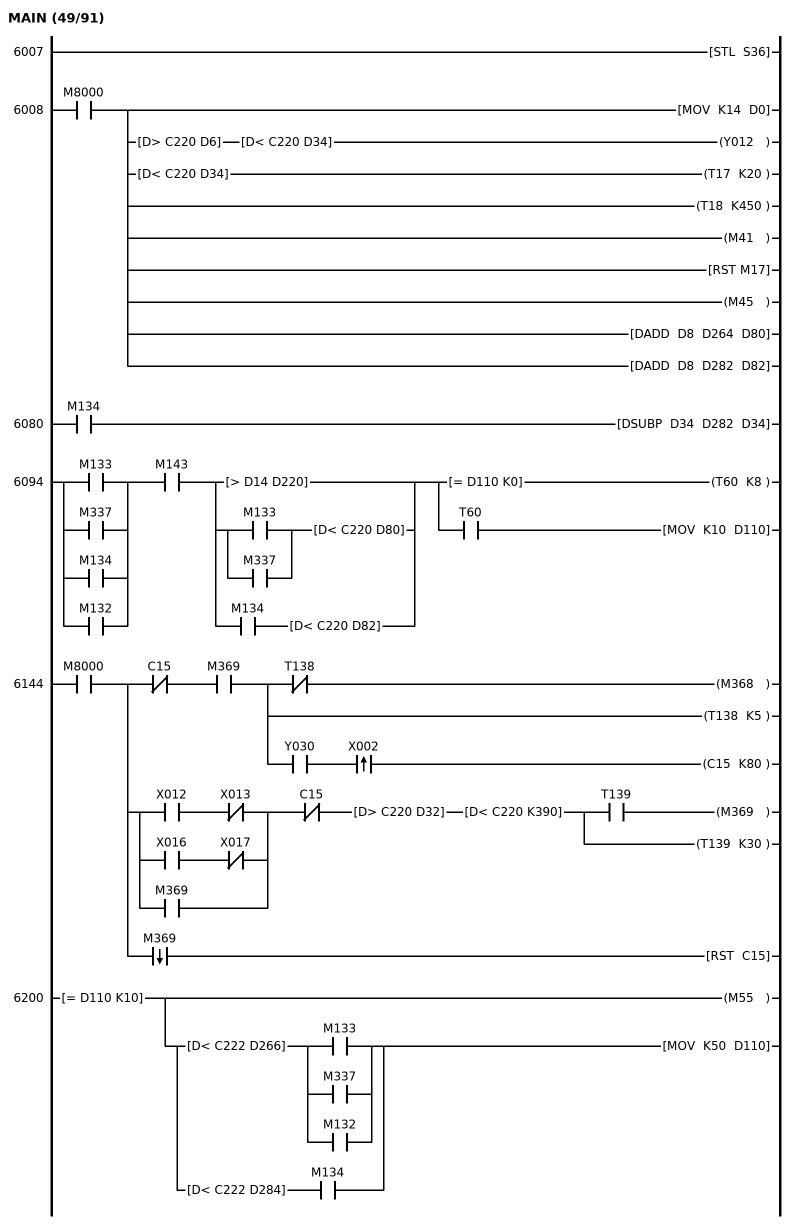
[picture p48: ladder of MAIN, rungs at steps 6007 to 6200]
6007  STL     S36
6008  LD      M8000
      MOV     K14 D0
      MPS
      ANDD>   C220 D6
      ANDD<   C220 D34
      OUT     Y012
      MRD
      ANDD<   C220 D34
      OUT     T17 K20
      MPP
      OUT     T18 K450
      OUT     M41
      RST     M17
      OUT     M45
      DADD    D8 D264 D80
      DADD    D8 D282 D82
6080  LD      M134
      DSUBP   D34 D282 D34
6094  LD      M133
      OR      M337
      OR      M134
      OR      M132
      AND     M143
      LD>     D14 D220
      LD      M133
      OR      M337
      ANDD<   C220 D80
      ORB
      LD      M134
      ANDD<   C220 D82
      ORB
      ANB
      MPS
      AND=    D110 K0
      OUT     T60 K8
      MPP
      AND     T60
      MOV     K10 D110
6144  LD      M8000
      MPS
      ANI     C15
      AND     M369
      MPS
      ANI     T138
      OUT     M368
      MPP
      OUT     T138 K5
      AND     Y030
      ANDP    X002
      OUT     C15 K80
      MRD
      LD      X012
      ANI     X013
      LD      X016
      ANI     X017
      ORB
      OR      M369
      ANB
      ANI     C15
      ANDD>   C220 D32
      ANDD<   C220 K390
      MPS
      AND     T139
      OUT     M369
      MPP
      OUT     T139 K30
      MPP
      ANDF    M369
      RST     C15
6200  LD=     D110 K10
      OUT     M55
      LDD<    C222 D266
      LD      M133
      OR      M337
      OR      M132
      ANB
      LDD<    C222 D284
      AND     M134
      ORB
      ANB
      MOV     K50 D110
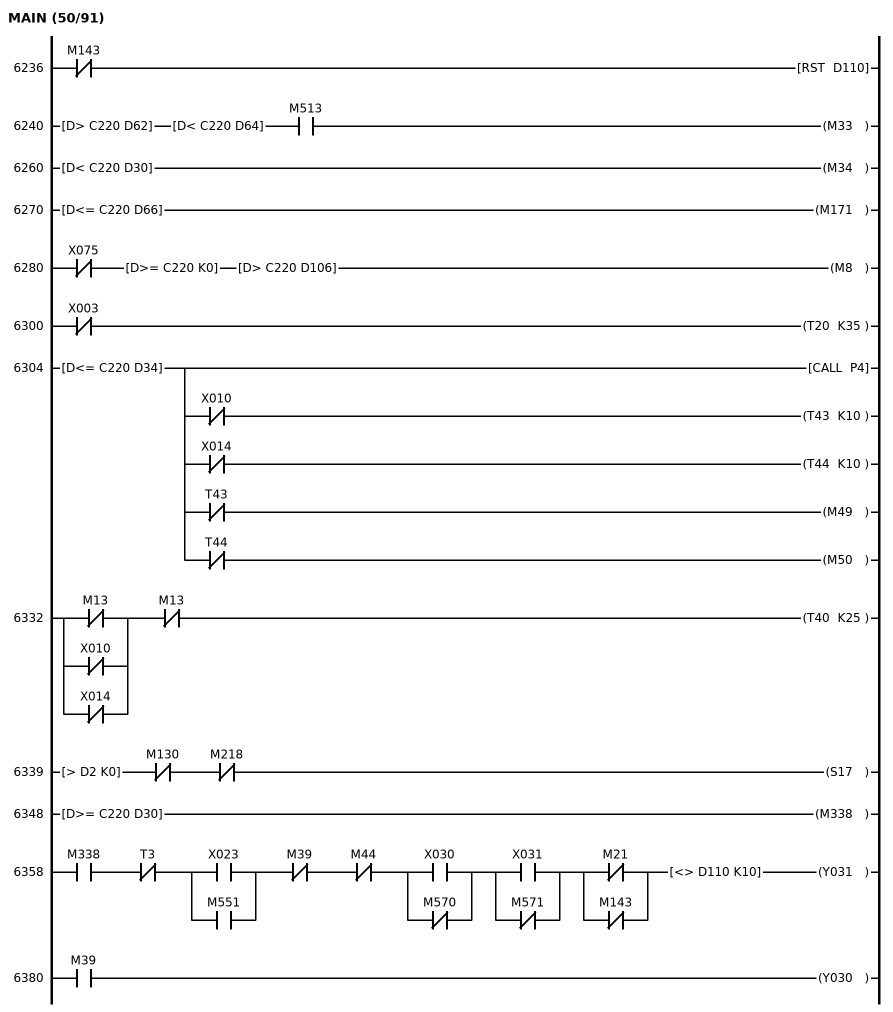
6236  LDI     M143
      RST     D110
6240  LDD>    C220 D62
      ANDD<   C220 D64
      AND     M513
      OUT     M33
6260  LDD<    C220 D30
      OUT     M34
6270  LDD<=   C220 D66
      OUT     M171
6280  LDI     X075
      ANDD>=  C220 K0
      ANDD>   C220 D106
      OUT     M8
6300  LDI     X003
      OUT     T20 K35
6304  LDD<=   C220 D34
      CALL    P4
      MPS
      ANI     X010
      OUT     T43 K10
      MRD
      ANI     X014
      OUT     T44 K10
      MRD
      ANI     T43
      OUT     M49
      MPP
      ANI     T44
      OUT     M50
6332  LDI     M13
      ORI     X010
      ORI     X014
      ANI     M13
      OUT     T40 K25
6339  LD>     D2 K0
      ANI     M130
      ANI     M218
      OUT     S17
6348  LDD>=   C220 D30
      OUT     M338
6358  LD      M338
      ANI     T3
      LD      X023
      OR      M551
      ANB
      ANI     M39
      ANI     M44
      LD      X030
      ORI     M570
      ANB
      LD      X031
      ORI     M571
      ANB
      LDI     M21
      ORI     M143
      ANB
      AND<>   D110 K10
      OUT     Y031
6380  LD      M39
      OUT     Y030
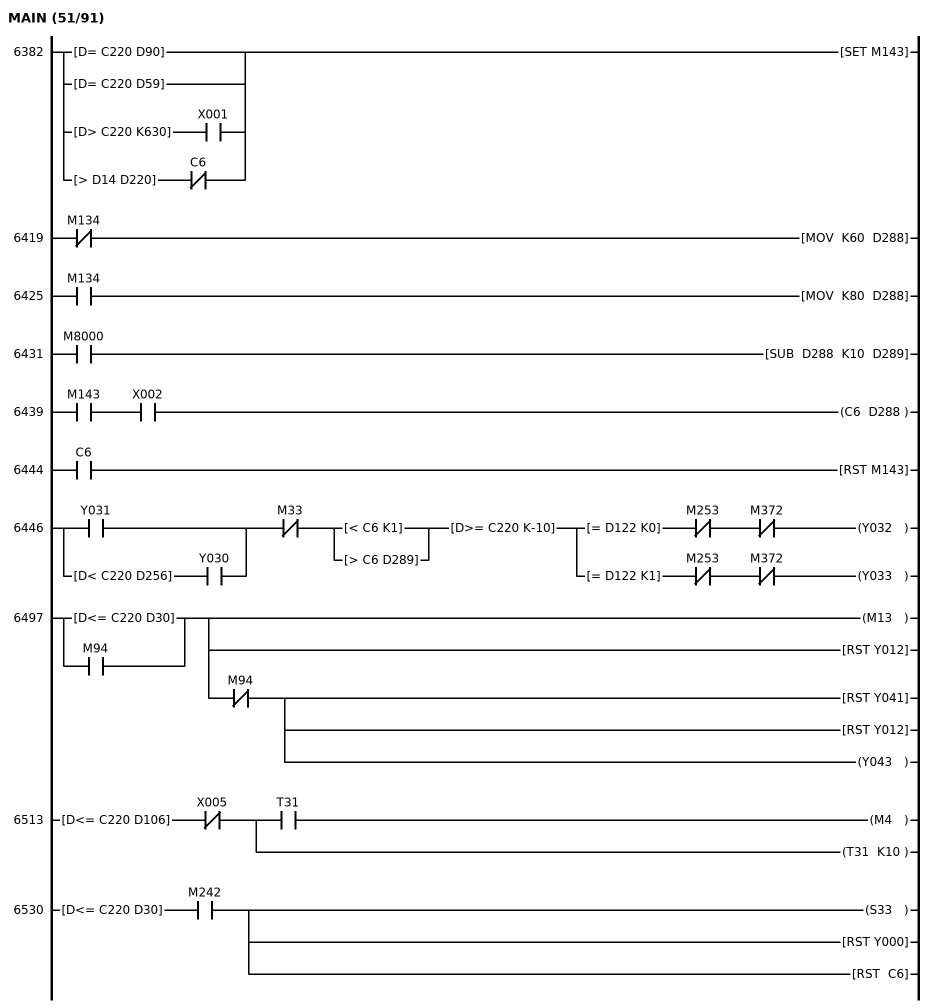
6382  LDD=    C220 D90
      ORD=    C220 D59
      LDD>    C220 K630
      AND     X001
      ORB
      LD>     D14 D220
      ANI     C6
      ORB
      SET     M143
6419  LDI     M134
      MOV     K60 D288
6425  LD      M134
      MOV     K80 D288
6431  LD      M8000
      SUB     D288 K10 D289
6439  LD      M143
      AND     X002
      OUT     C6 D288
6444  LD      C6
      RST     M143
6446  LD      Y031
      LDD<    C220 D256
      AND     Y030
      ORB
      ANI     M33
      LD<     C6 K1
      OR>     C6 D289
      ANB
      ANDD>=  C220 K-10
      MPS
      AND=    D122 K0
      ANI     M253
      ANI     M372
      OUT     Y032
      MPP
      AND=    D122 K1
      ANI     M253
      ANI     M372
      OUT     Y033
6497  LDD<=   C220 D30
      OR      M94
      OUT     M13
      RST     Y012
      ANI     M94
      RST     Y041
      RST     Y012
      OUT     Y043
6513  LDD<=   C220 D106
      ANI     X005
      MPS
      AND     T31
      OUT     M4
      MPP
      OUT     T31 K10
6530  LDD<=   C220 D30
      AND     M242
      OUT     S33
      RST     Y000
      RST     C6
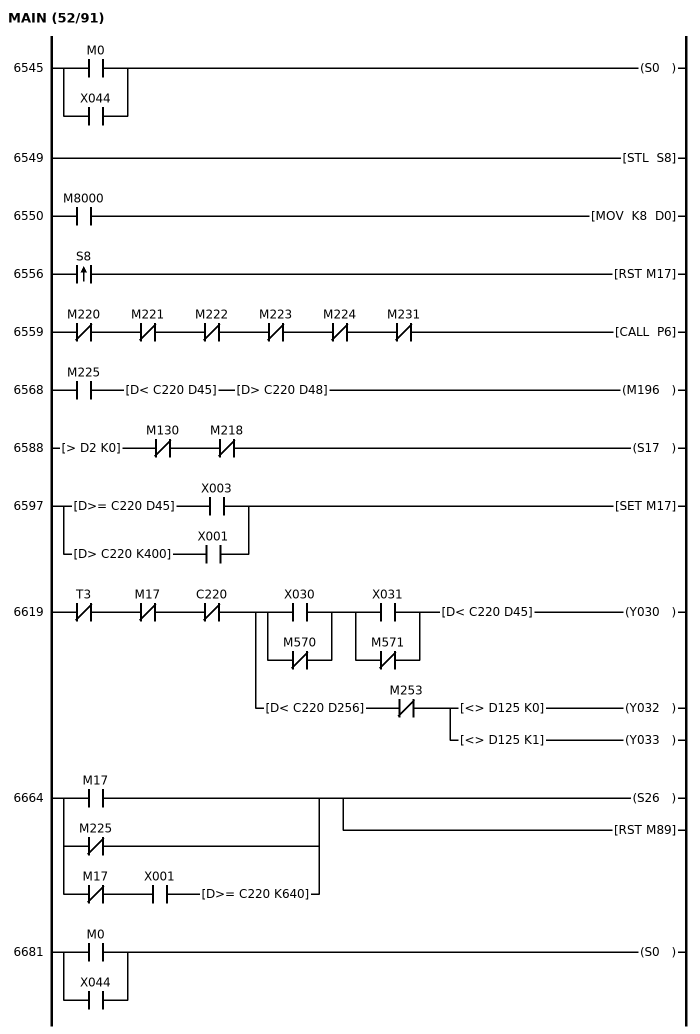
6545  LD      M0
      OR      X044
      OUT     S0
6549  STL     S8
6550  LD      M8000
      MOV     K8 D0
6556  LDP     S8
      RST     M17
6559  LDI     M220
      ANI     M221
      ANI     M222
      ANI     M223
      ANI     M224
      ANI     M231
      CALL    P6
6568  LD      M225
      ANDD<   C220 D45
      ANDD>   C220 D48
      OUT     M196
6588  LD>     D2 K0
      ANI     M130
      ANI     M218
      OUT     S17
6597  LDD>=   C220 D45
      AND     X003
      LDD>    C220 K400
      AND     X001
      ORB
      SET     M17
6619  LDI     T3
      ANI     M17
      ANI     C220
      MPS
      LD      X030
      ORI     M570
      ANB
      LD      X031
      ORI     M571
      ANB
      ANDD<   C220 D45
      OUT     Y030
      MPP
      ANDD<   C220 D256
      ANI     M253
      MPS
      AND<>   D125 K0
      OUT     Y032
      MPP
      AND<>   D125 K1
      OUT     Y033
6664  LD      M17
      ORI     M225
      LDI     M17
      AND     X001
      ANDD>=  C220 K640
      ORB
      OUT     S26
      RST     M89
6681  LD      M0
      OR      X044
      OUT     S0
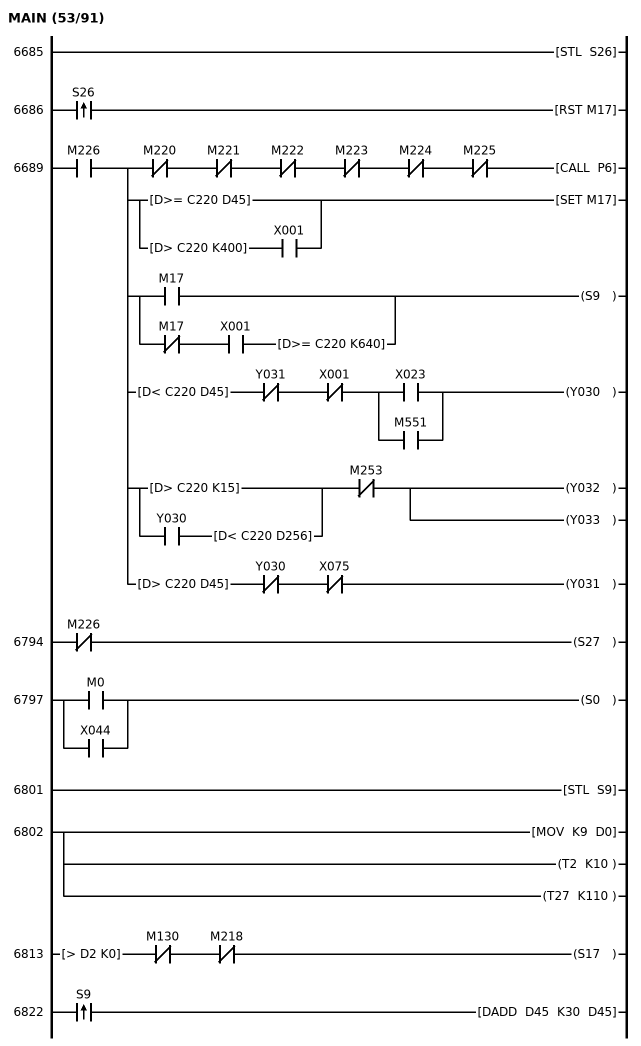
6685  STL     S26
6686  LDP     S26
      RST     M17
6689  LD      M226
      MPS
      ANI     M220
      ANI     M221
      ANI     M222
      ANI     M223
      ANI     M224
      ANI     M225
      CALL    P6
      MRD
      LDD>=   C220 D45
      LDD>    C220 K400
      AND     X001
      ORB
      ANB
      SET     M17
      MRD
      LD      M17
      LDI     M17
      AND     X001
      ANDD>=  C220 K640
      ORB
      ANB
      OUT     S9
      MRD
      ANDD<   C220 D45
      ANI     Y031
      ANI     X001
      LD      X023
      OR      M551
      ANB
      OUT     Y030
      MRD
      LDD>    C220 K15
      LD      Y030
      ANDD<   C220 D256
      ORB
      ANB
      ANI     M253
      OUT     Y032
      OUT     Y033
      MPP
      ANDD>   C220 D45
      ANI     Y030
      ANI     X075
      OUT     Y031
6794  LDI     M226
      OUT     S27
6797  LD      M0
      OR      X044
      OUT     S0
6801  STL     S9
6802  MOV     K9 D0
      OUT     T2 K10
      OUT     T27 K110
6813  LD>     D2 K0
      ANI     M130
      ANI     M218
      OUT     S17
6822  LDP     S9
      DADD    D45 K30 D45
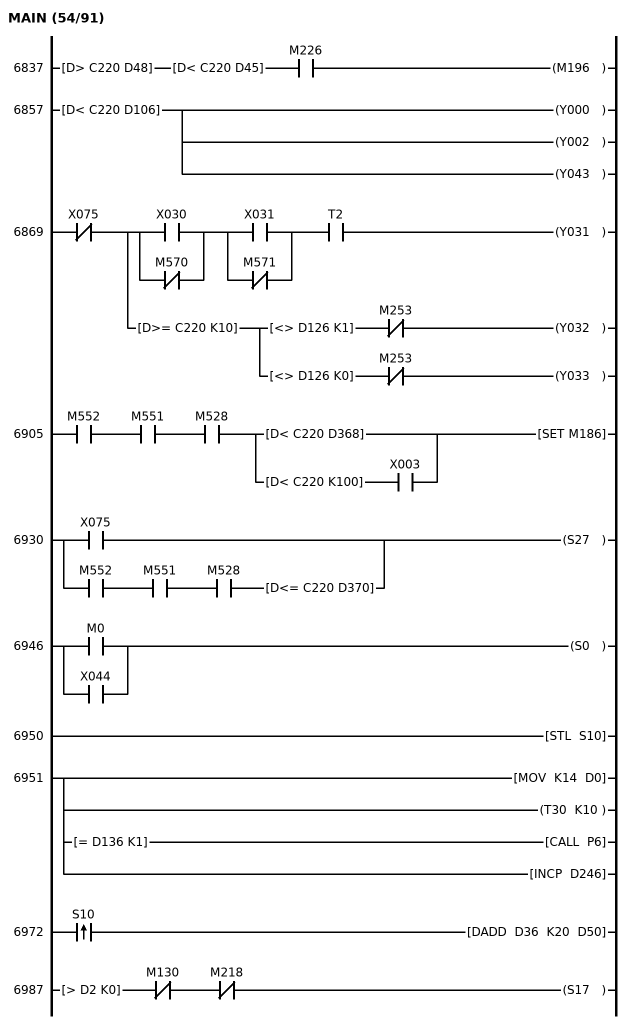
6837  LDD>    C220 D48
      ANDD<   C220 D45
      AND     M226
      OUT     M196
6857  LDD<    C220 D106
      OUT     Y000
      OUT     Y002
      OUT     Y043
6869  LDI     X075
      MPS
      LD      X030
      ORI     M570
      ANB
      LD      X031
      ORI     M571
      ANB
      AND     T2
      OUT     Y031
      MPP
      ANDD>=  C220 K10
      MPS
      AND<>   D126 K1
      ANI     M253
      OUT     Y032
      MPP
      AND<>   D126 K0
      ANI     M253
      OUT     Y033
6905  LD      M552
      AND     M551
      AND     M528
      LDD<    C220 D368
      LDD<    C220 K100
      AND     X003
      ORB
      ANB
      SET     M186
6930  LD      X075
      LD      M552
      AND     M551
      AND     M528
      ANDD<=  C220 D370
      ORB
      OUT     S27
6946  LD      M0
      OR      X044
      OUT     S0
6950  STL     S10
6951  MOV     K14 D0
      OUT     T30 K10
      MPS
      AND=    D136 K1
      CALL    P6
      MPP
      INCP    D246
6972  LDP     S10
      DADD    D36 K20 D50
6987  LD>     D2 K0
      ANI     M130
      ANI     M218
      OUT     S17
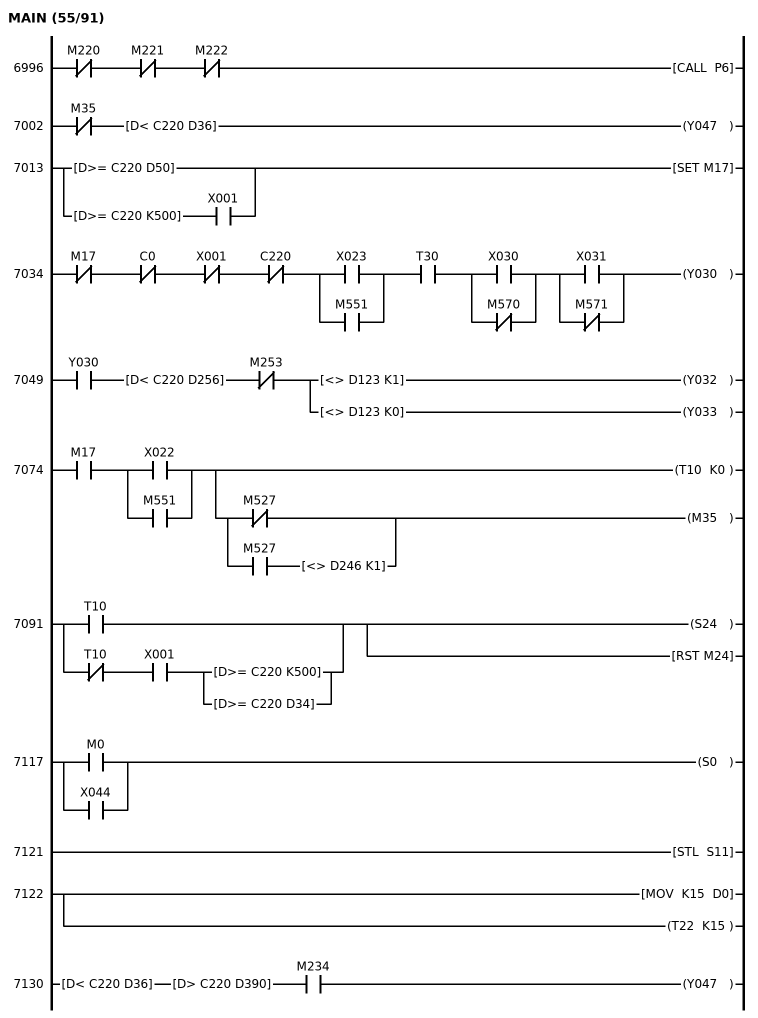
6996  LDI     M220
      ANI     M221
      ANI     M222
      CALL    P6
7002  LDI     M35
      ANDD<   C220 D36
      OUT     Y047
7013  LDD>=   C220 D50
      LDD>=   C220 K500
      AND     X001
      ORB
      SET     M17
7034  LDI     M17
      ANI     C0
      ANI     X001
      ANI     C220
      LD      X023
      OR      M551
      ANB
      AND     T30
      LD      X030
      ORI     M570
      ANB
      LD      X031
      ORI     M571
      ANB
      OUT     Y030
7049  LD      Y030
      ANDD<   C220 D256
      ANI     M253
      MPS
      AND<>   D123 K1
      OUT     Y032
      MPP
      AND<>   D123 K0
      OUT     Y033
7074  LD      M17
      LD      X022
      OR      M551
      ANB
      OUT     T10 K0
      LDI     M527
      LD      M527
      AND<>   D246 K1
      ORB
      ANB
      OUT     M35
7091  LD      T10
      LDI     T10
      AND     X001
      LDD>=   C220 K500
      ORD>=   C220 D34
      ANB
      ORB
      OUT     S24
      RST     M24
7117  LD      M0
      OR      X044
      OUT     S0
7121  STL     S11
7122  MOV     K15 D0
      OUT     T22 K15
7130  LDD<    C220 D36
      ANDD>   C220 D390
      AND     M234
      OUT     Y047
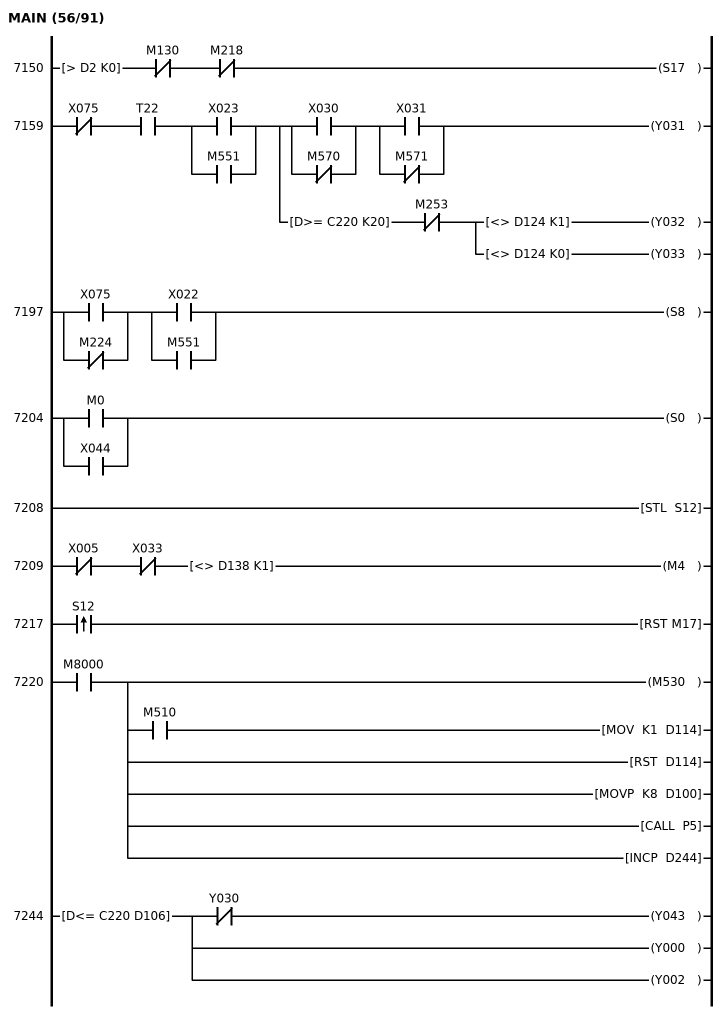
7150  LD>     D2 K0
      ANI     M130
      ANI     M218
      OUT     S17
7159  LDI     X075
      AND     T22
      LD      X023
      OR      M551
      ANB
      MPS
      LD      X030
      ORI     M570
      ANB
      LD      X031
      ORI     M571
      ANB
      OUT     Y031
      MPP
      ANDD>=  C220 K20
      ANI     M253
      MPS
      AND<>   D124 K1
      OUT     Y032
      MPP
      AND<>   D124 K0
      OUT     Y033
7197  LD      X075
      ORI     M224
      LD      X022
      OR      M551
      ANB
      OUT     S8
7204  LD      M0
      OR      X044
      OUT     S0
7208  STL     S12
7209  LDI     X005
      ANI     X033
      AND<>   D138 K1
      OUT     M4
7217  LDP     S12
      RST     M17
7220  LD      M8000
      OUT     M530
      MPS
      AND     M510
      MOV     K1 D114
      MPP
      RST     D114
      MOVP    K8 D100
      CALL    P5
      INCP    D244
7244  LDD<=   C220 D106
      MPS
      ANI     Y030
      OUT     Y043
      MPP
      OUT     Y000
      OUT     Y002
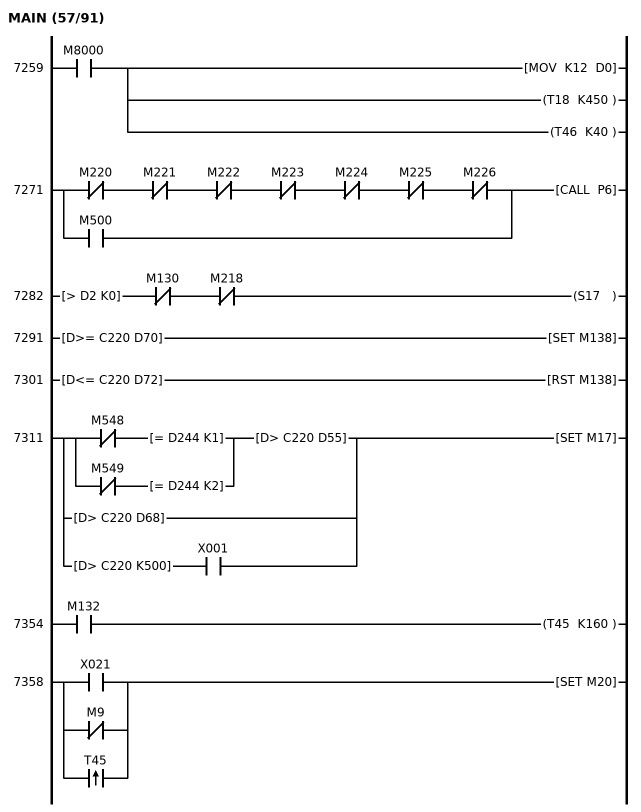
7259  LD      M8000
      MOV     K12 D0
      OUT     T18 K450
      OUT     T46 K40
7271  LDI     M220
      ANI     M221
      ANI     M222
      ANI     M223
      ANI     M224
      ANI     M225
      ANI     M226
      OR      M500
      CALL    P6
7282  LD>     D2 K0
      ANI     M130
      ANI     M218
      OUT     S17
7291  LDD>=   C220 D70
      SET     M138
7301  LDD<=   C220 D72
      RST     M138
7311  LDI     M548
      AND=    D244 K1
      LDI     M549
      AND=    D244 K2
      ORB
      ANDD>   C220 D55
      ORD>    C220 D68
      LDD>    C220 K500
      AND     X001
      ORB
      SET     M17
7354  LD      M132
      OUT     T45 K160
7358  LD      X021
      ORI     M9
      ORP     T45
      SET     M20
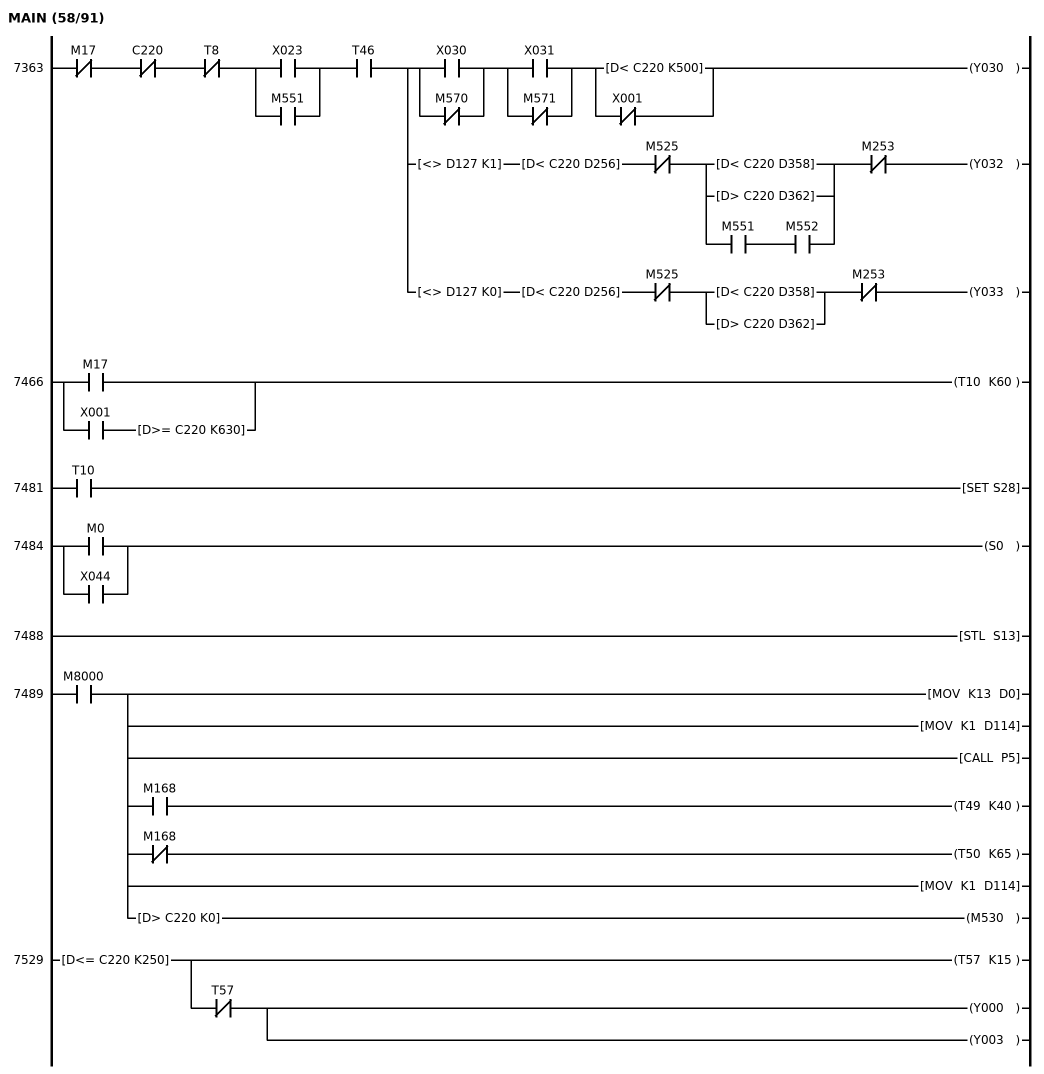
7363  LDI     M17
      ANI     C220
      ANI     T8
      LD      X023
      OR      M551
      ANB
      AND     T46
      MPS
      LD      X030
      ORI     M570
      ANB
      LD      X031
      ORI     M571
      ANB
      LDD<    C220 K500
      ORI     X001
      ANB
      OUT     Y030
      MRD
      AND<>   D127 K1
      ANDD<   C220 D256
      ANI     M525
      LDD<    C220 D358
      ORD>    C220 D362
      LD      M551
      AND     M552
      ORB
      ANB
      ANI     M253
      OUT     Y032
      MPP
      AND<>   D127 K0
      ANDD<   C220 D256
      ANI     M525
      LDD<    C220 D358
      ORD>    C220 D362
      ANB
      ANI     M253
      OUT     Y033
7466  LD      M17
      LD      X001
      ANDD>=  C220 K630
      ORB
      OUT     T10 K60
7481  LD      T10
      SET     S28
7484  LD      M0
      OR      X044
      OUT     S0
7488  STL     S13
7489  LD      M8000
      MOV     K13 D0
      MOV     K1 D114
      CALL    P5
      MPS
      AND     M168
      OUT     T49 K40
      MRD
      ANI     M168
      OUT     T50 K65
      MPP
      MOV     K1 D114
      ANDD>   C220 K0
      OUT     M530
7529  LDD<=   C220 K250
      OUT     T57 K15
      ANI     T57
      OUT     Y000
      OUT     Y003
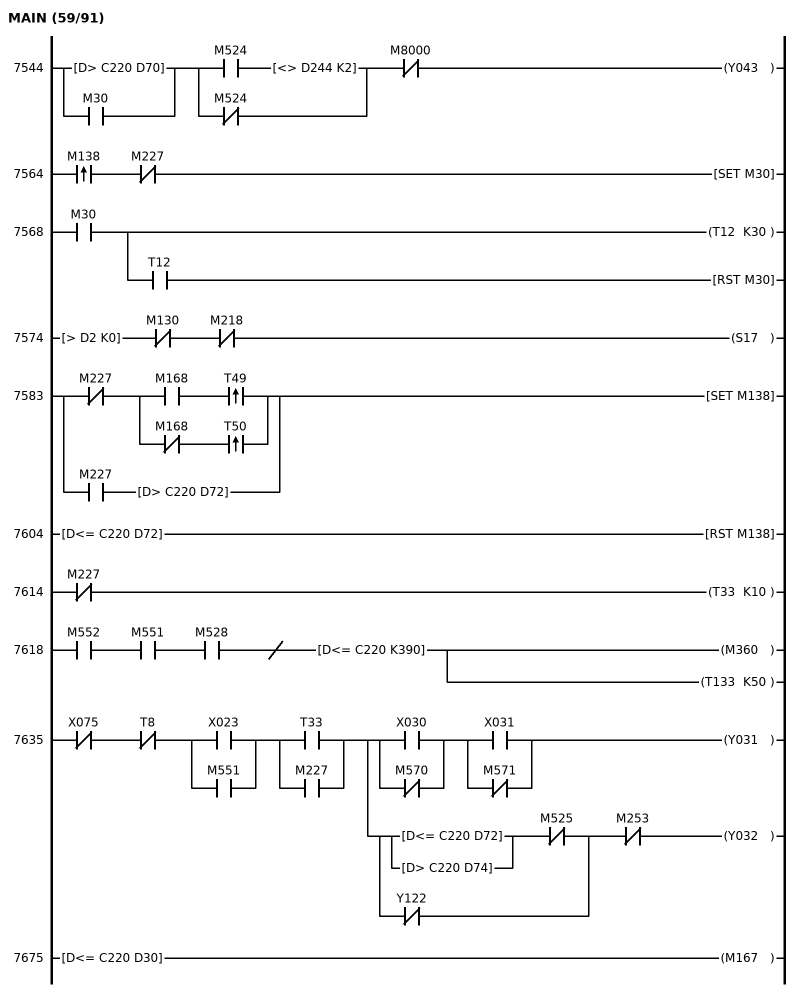
7544  LDD>    C220 D70
      OR      M30
      LD      M524
      AND<>   D244 K2
      ORI     M524
      ANB
      ANI     M8000
      OUT     Y043
7564  LDP     M138
      ANI     M227
      SET     M30
7568  LD      M30
      OUT     T12 K30
      AND     T12
      RST     M30
7574  LD>     D2 K0
      ANI     M130
      ANI     M218
      OUT     S17
7583  LDI     M227
      LD      M168
      ANDP    T49
      LDI     M168
      ANDP    T50
      ORB
      ANB
      LD      M227
      ANDD>   C220 D72
      ORB
      SET     M138
7604  LDD<=   C220 D72
      RST     M138
7614  LDI     M227
      OUT     T33 K10
7618  LD      M552
      AND     M551
      AND     M528
      INV
      ANDD<=  C220 K390
      OUT     M360
      OUT     T133 K50
7635  LDI     X075
      ANI     T8
      LD      X023
      OR      M551
      ANB
      LD      T33
      OR      M227
      ANB
      MPS
      LD      X030
      ORI     M570
      ANB
      LD      X031
      ORI     M571
      ANB
      OUT     Y031
      MPP
      LDD<=   C220 D72
      ORD>    C220 D74
      ANI     M525
      ORI     Y122
      ANB
      ANI     M253
      OUT     Y032
7675  LDD<=   C220 D30
      OUT     M167
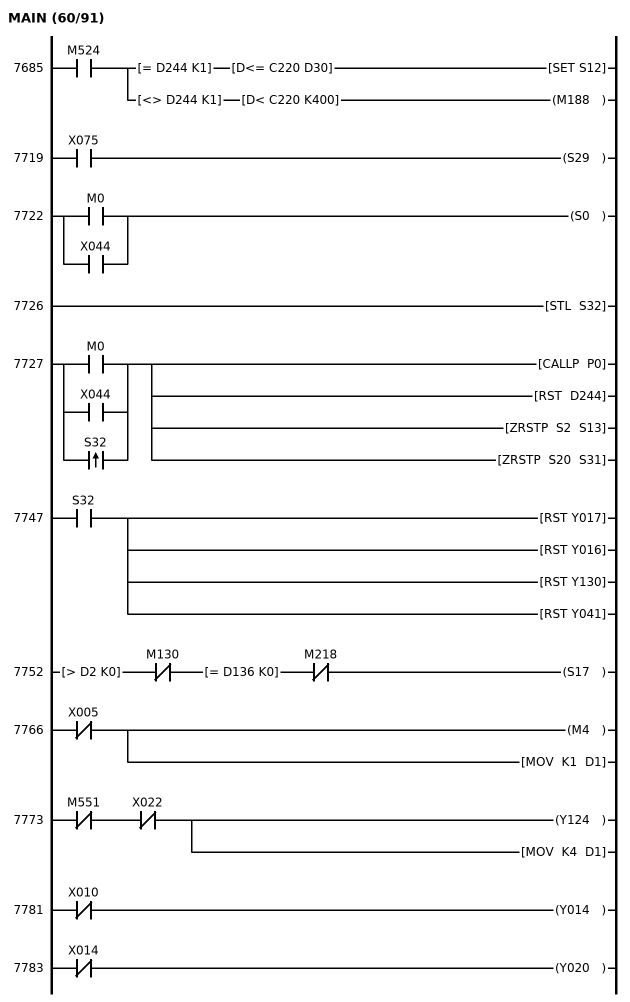
7685  LD      M524
      MPS
      AND=    D244 K1
      ANDD<=  C220 D30
      SET     S12
      MPP
      AND<>   D244 K1
      ANDD<   C220 K400
      OUT     M188
7719  LD      X075
      OUT     S29
7722  LD      M0
      OR      X044
      OUT     S0
7726  STL     S32
7727  LD      M0
      OR      X044
      ORP     S32
      CALLP   P0
      RST     D244
      ZRSTP   S2 S13
      ZRSTP   S20 S31
7747  LD      S32
      RST     Y017
      RST     Y016
      RST     Y130
      RST     Y041
7752  LD>     D2 K0
      ANI     M130
      AND=    D136 K0
      ANI     M218
      OUT     S17
7766  LDI     X005
      OUT     M4
      MOV     K1 D1
7773  LDI     M551
      ANI     X022
      OUT     Y124
      MOV     K4 D1
7781  LDI     X010
      OUT     Y014
7783  LDI     X014
      OUT     Y020
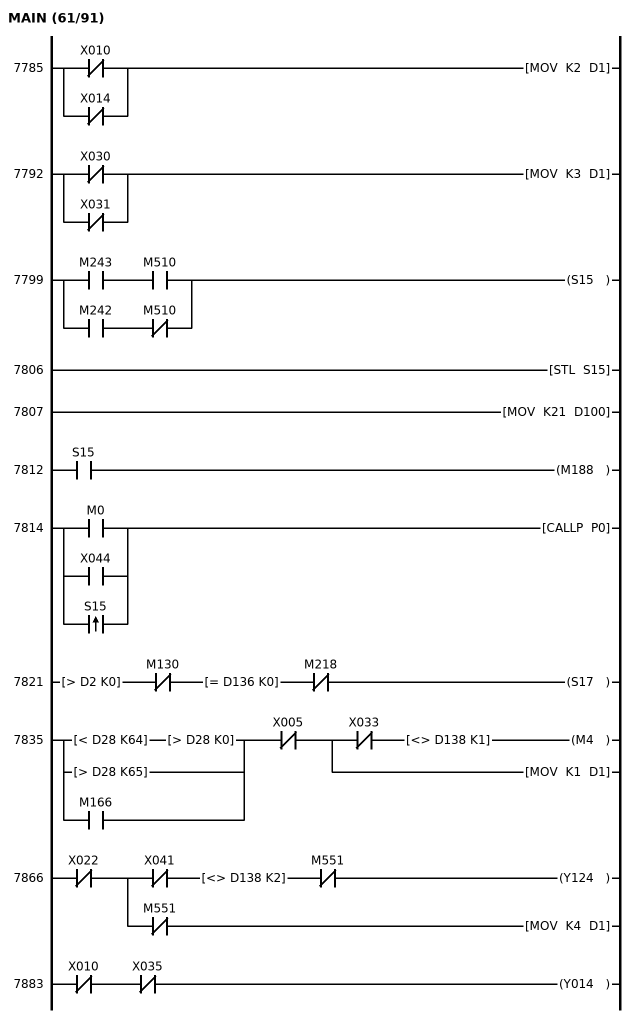
7785  LDI     X010
      ORI     X014
      MOV     K2 D1
7792  LDI     X030
      ORI     X031
      MOV     K3 D1
7799  LD      M243
      AND     M510
      LD      M242
      ANI     M510
      ORB
      OUT     S15
7806  STL     S15
7807  MOV     K21 D100
7812  LD      S15
      OUT     M188
7814  LD      M0
      OR      X044
      ORP     S15
      CALLP   P0
7821  LD>     D2 K0
      ANI     M130
      AND=    D136 K0
      ANI     M218
      OUT     S17
7835  LD<     D28 K64
      AND>    D28 K0
      OR>     D28 K65
      OR      M166
      ANI     X005
      MPS
      ANI     X033
      AND<>   D138 K1
      OUT     M4
      MPP
      MOV     K1 D1
7866  LDI     X022
      MPS
      ANI     X041
      AND<>   D138 K2
      ANI     M551
      OUT     Y124
      MPP
      ANI     M551
      MOV     K4 D1
7883  LDI     X010
      ANI     X035
      OUT     Y014
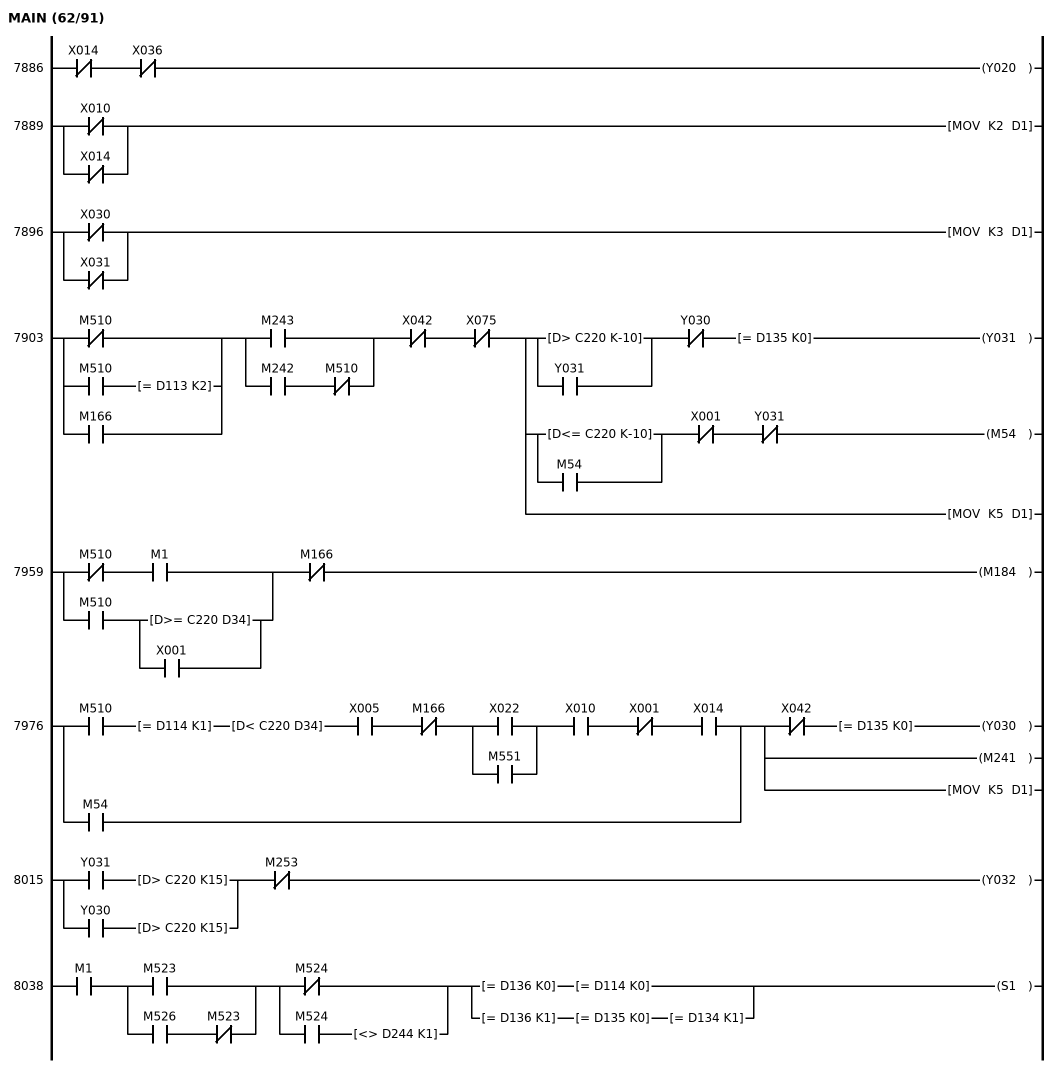
7886  LDI     X014
      ANI     X036
      OUT     Y020
7889  LDI     X010
      ORI     X014
      MOV     K2 D1
7896  LDI     X030
      ORI     X031
      MOV     K3 D1
7903  LDI     M510
      LD      M510
      AND=    D113 K2
      ORB
      OR      M166
      LD      M243
      LD      M242
      ANI     M510
      ORB
      ANB
      ANI     X042
      ANI     X075
      MPS
      LDD>    C220 K-10
      OR      Y031
      ANB
      ANI     Y030
      AND=    D135 K0
      OUT     Y031
      MRD
      LDD<=   C220 K-10
      OR      M54
      ANB
      ANI     X001
      ANI     Y031
      OUT     M54
      MPP
      MOV     K5 D1
7959  LDI     M510
      AND     M1
      LD      M510
      LDD>=   C220 D34
      OR      X001
      ANB
      ORB
      ANI     M166
      OUT     M184
7976  LD      M510
      AND=    D114 K1
      ANDD<   C220 D34
      AND     X005
      ANI     M166
      LD      X022
      OR      M551
      ANB
      AND     X010
      ANI     X001
      AND     X014
      OR      M54
      MPS
      ANI     X042
      AND=    D135 K0
      OUT     Y030
      MPP
      OUT     M241
      MOV     K5 D1
8015  LD      Y031
      ANDD>   C220 K15
      LD      Y030
      ANDD>   C220 K15
      ORB
      ANI     M253
      OUT     Y032
8038  LD      M1
      LD      M523
      LD      M526
      ANI     M523
      ORB
      ANB
      LDI     M524
      LD      M524
      AND<>   D244 K1
      ORB
      ANB
      LD=     D136 K0
      AND=    D114 K0
      LD=     D136 K1
      AND=    D135 K0
      AND=    D134 K1
      ORB
      ANB
      OUT     S1
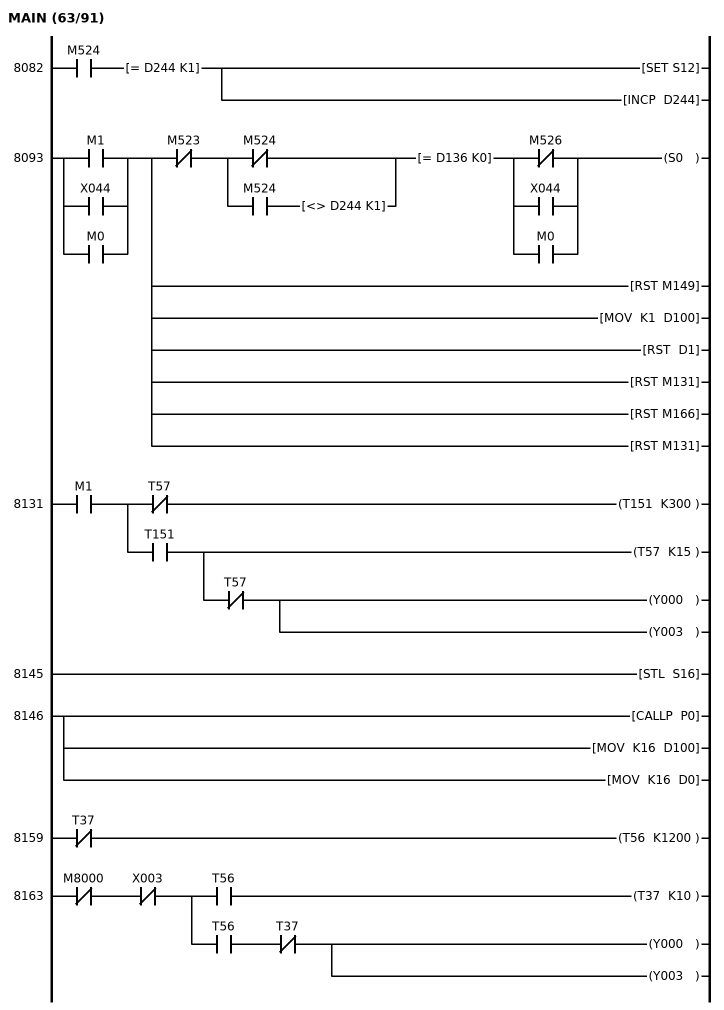
8082  LD      M524
      AND=    D244 K1
      SET     S12
      INCP    D244
8093  LD      M1
      OR      X044
      OR      M0
      MPS
      ANI     M523
      LDI     M524
      LD      M524
      AND<>   D244 K1
      ORB
      ANB
      AND=    D136 K0
      LDI     M526
      OR      X044
      OR      M0
      ANB
      OUT     S0
      MPP
      RST     M149
      MOV     K1 D100
      RST     D1
      RST     M131
      RST     M166
      RST     M131
8131  LD      M1
      MPS
      ANI     T57
      OUT     T151 K300
      MPP
      AND     T151
      OUT     T57 K15
      ANI     T57
      OUT     Y000
      OUT     Y003
8145  STL     S16
8146  CALLP   P0
      MOV     K16 D100
      MOV     K16 D0
8159  LDI     T37
      OUT     T56 K1200
8163  LDI     M8000
      ANI     X003
      MPS
      AND     T56
      OUT     T37 K10
      MPP
      AND     T56
      ANI     T37
      OUT     Y000
      OUT     Y003
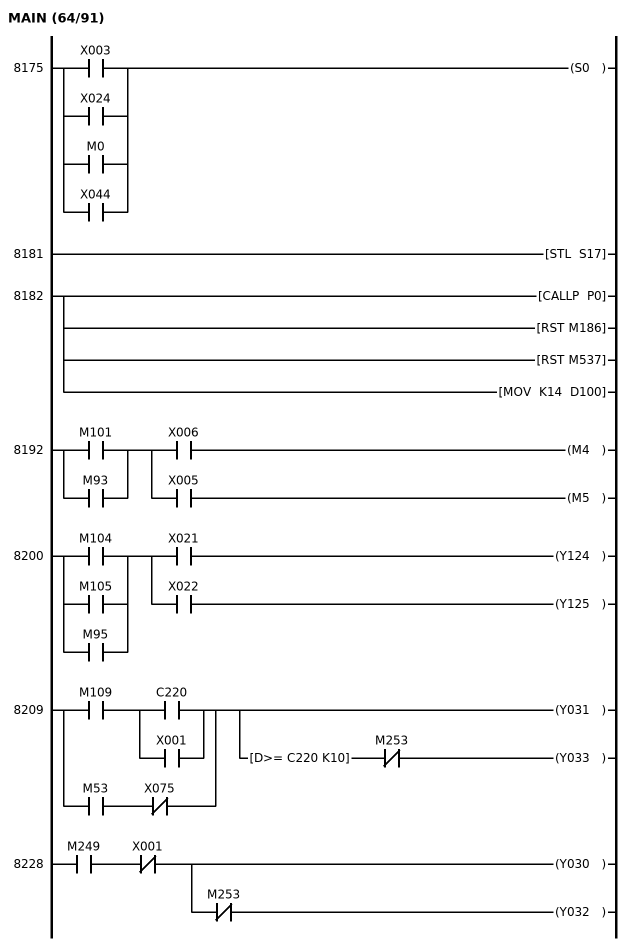
8175  LD      X003
      OR      X024
      OR      M0
      OR      X044
      OUT     S0
8181  STL     S17
8182  CALLP   P0
      RST     M186
      RST     M537
      MOV     K14 D100
8192  LD      M101
      OR      M93
      MPS
      AND     X006
      OUT     M4
      MPP
      AND     X005
      OUT     M5
8200  LD      M104
      OR      M105
      OR      M95
      MPS
      AND     X021
      OUT     Y124
      MPP
      AND     X022
      OUT     Y125
8209  LD      M109
      LD      C220
      OR      X001
      ANB
      LD      M53
      ANI     X075
      ORB
      OUT     Y031
      ANDD>=  C220 K10
      ANI     M253
      OUT     Y033
8228  LD      M249
      ANI     X001
      OUT     Y030
      ANI     M253
      OUT     Y032
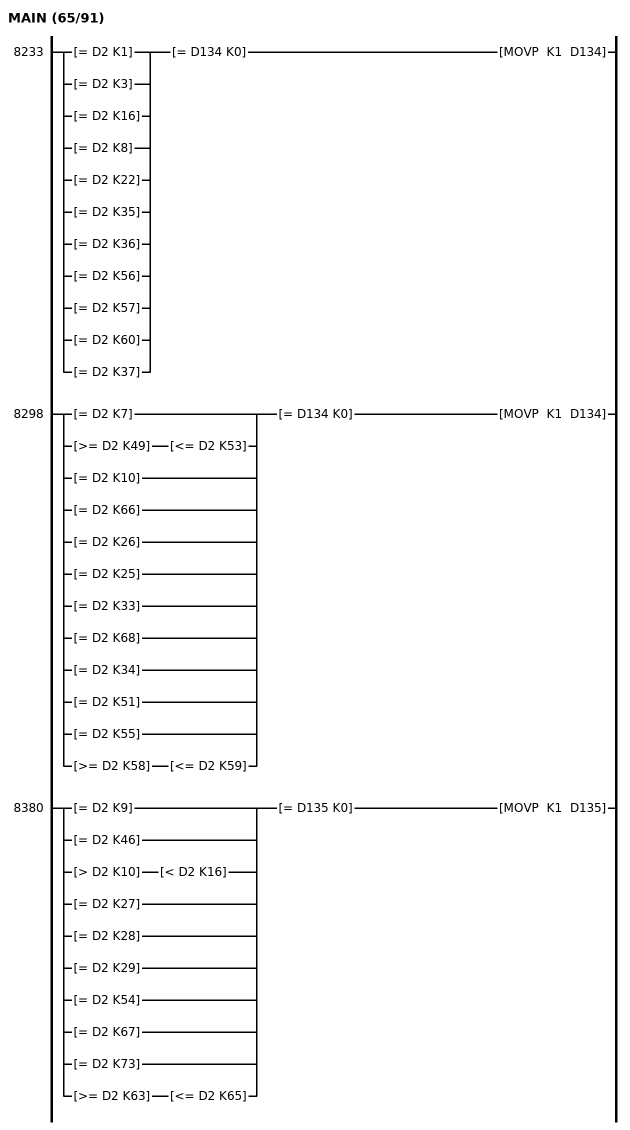
8233  LD=     D2 K1
      OR=     D2 K3
      OR=     D2 K16
      OR=     D2 K8
      OR=     D2 K22
      OR=     D2 K35
      OR=     D2 K36
      OR=     D2 K56
      OR=     D2 K57
      OR=     D2 K60
      OR=     D2 K37
      AND=    D134 K0
      MOVP    K1 D134
8298  LD=     D2 K7
      LD>=    D2 K49
      AND<=   D2 K53
      ORB
      OR=     D2 K10
      OR=     D2 K66
      OR=     D2 K26
      OR=     D2 K25
      OR=     D2 K33
      OR=     D2 K68
      OR=     D2 K34
      OR=     D2 K51
      OR=     D2 K55
      LD>=    D2 K58
      AND<=   D2 K59
      ORB
      AND=    D134 K0
      MOVP    K1 D134
8380  LD=     D2 K9
      OR=     D2 K46
      LD>     D2 K10
      AND<    D2 K16
      ORB
      OR=     D2 K27
      OR=     D2 K28
      OR=     D2 K29
      OR=     D2 K54
      OR=     D2 K67
      OR=     D2 K73
      LD>=    D2 K63
      AND<=   D2 K65
      ORB
      AND=    D135 K0
      MOVP    K1 D135
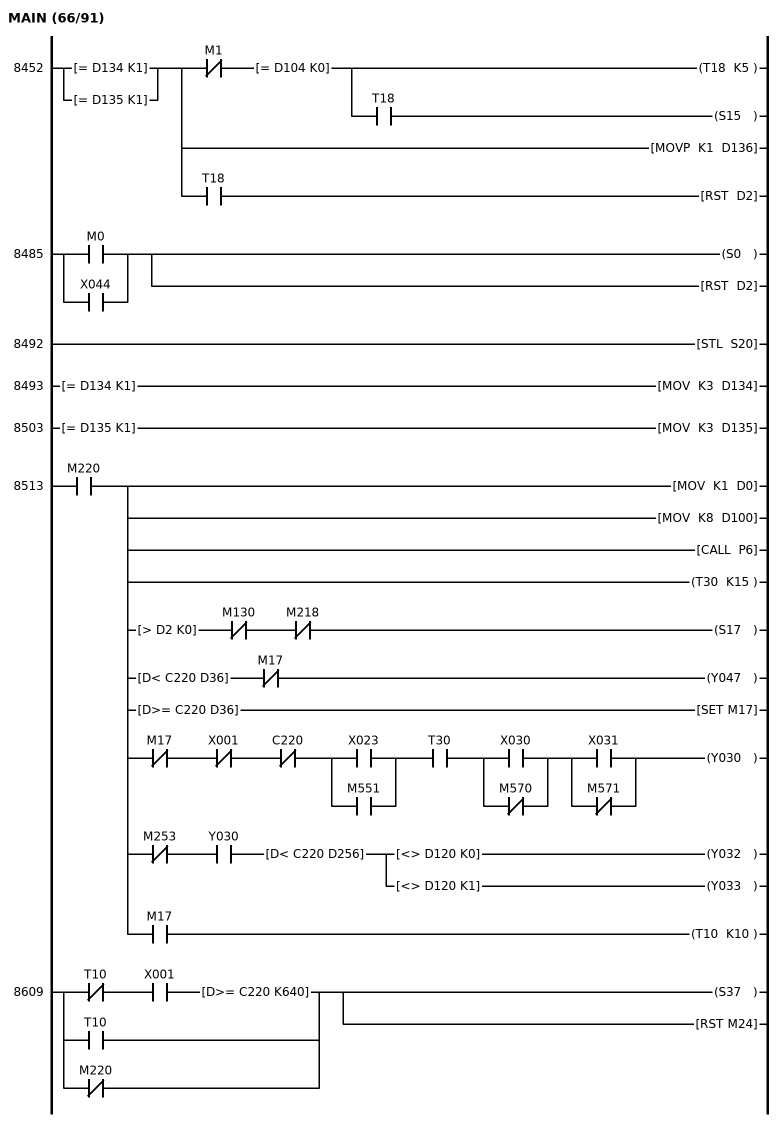
8452  LD=     D134 K1
      OR=     D135 K1
      MPS
      ANI     M1
      AND=    D104 K0
      OUT     T18 K5
      AND     T18
      OUT     S15
      MPP
      MOVP    K1 D136
      AND     T18
      RST     D2
8485  LD      M0
      OR      X044
      OUT     S0
      RST     D2
8492  STL     S20
8493  LD=     D134 K1
      MOV     K3 D134
8503  LD=     D135 K1
      MOV     K3 D135
8513  LD      M220
      MOV     K1 D0
      MOV     K8 D100
      CALL    P6
      OUT     T30 K15
      MPS
      AND>    D2 K0
      ANI     M130
      ANI     M218
      OUT     S17
      MRD
      ANDD<   C220 D36
      ANI     M17
      OUT     Y047
      MRD
      ANDD>=  C220 D36
      SET     M17
      MRD
      ANI     M17
      ANI     X001
      ANI     C220
      LD      X023
      OR      M551
      ANB
      AND     T30
      LD      X030
      ORI     M570
      ANB
      LD      X031
      ORI     M571
      ANB
      OUT     Y030
      MRD
      ANI     M253
      AND     Y030
      ANDD<   C220 D256
      MPS
      AND<>   D120 K0
      OUT     Y032
      MPP
      AND<>   D120 K1
      OUT     Y033
      MPP
      AND     M17
      OUT     T10 K10
8609  LDI     T10
      AND     X001
      ANDD>=  C220 K640
      OR      T10
      ORI     M220
      OUT     S37
      RST     M24
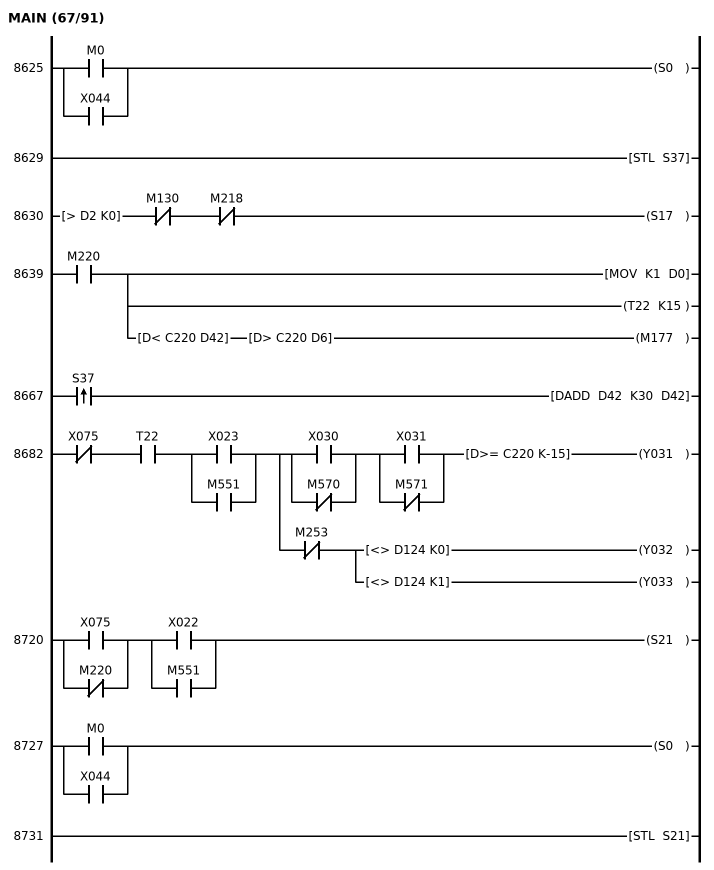
8625  LD      M0
      OR      X044
      OUT     S0
8629  STL     S37
8630  LD>     D2 K0
      ANI     M130
      ANI     M218
      OUT     S17
8639  LD      M220
      MOV     K1 D0
      OUT     T22 K15
      ANDD<   C220 D42
      ANDD>   C220 D6
      OUT     M177
8667  LDP     S37
      DADD    D42 K30 D42
8682  LDI     X075
      AND     T22
      LD      X023
      OR      M551
      ANB
      MPS
      LD      X030
      ORI     M570
      ANB
      LD      X031
      ORI     M571
      ANB
      ANDD>=  C220 K-15
      OUT     Y031
      MPP
      ANI     M253
      MPS
      AND<>   D124 K0
      OUT     Y032
      MPP
      AND<>   D124 K1
      OUT     Y033
8720  LD      X075
      ORI     M220
      LD      X022
      OR      M551
      ANB
      OUT     S21
8727  LD      M0
      OR      X044
      OUT     S0
8731  STL     S21
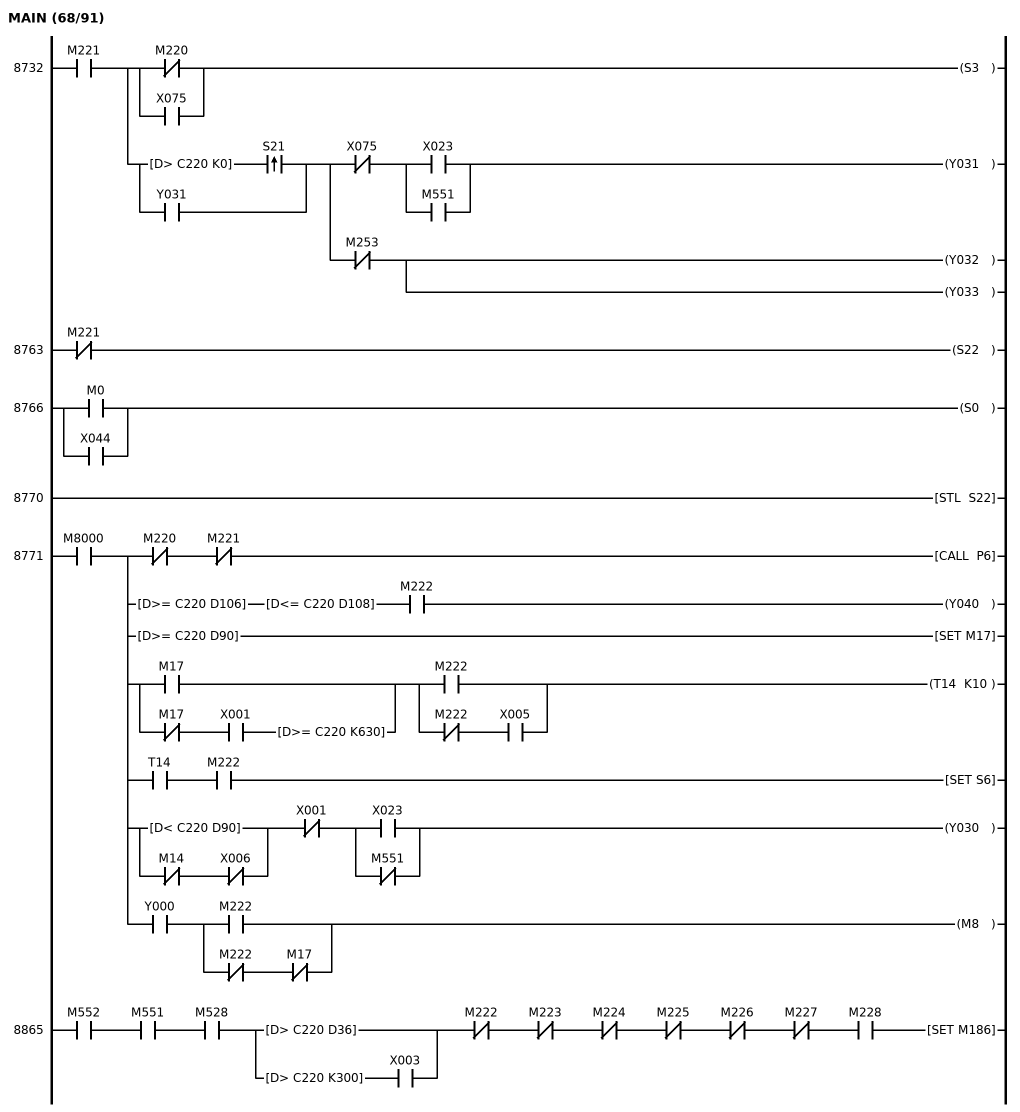
8732  LD      M221
      MPS
      LDI     M220
      OR      X075
      ANB
      OUT     S3
      MPP
      LDD>    C220 K0
      ANDP    S21
      OR      Y031
      ANB
      MPS
      ANI     X075
      LD      X023
      OR      M551
      ANB
      OUT     Y031
      MPP
      ANI     M253
      OUT     Y032
      OUT     Y033
8763  LDI     M221
      OUT     S22
8766  LD      M0
      OR      X044
      OUT     S0
8770  STL     S22
8771  LD      M8000
      MPS
      ANI     M220
      ANI     M221
      CALL    P6
      MRD
      ANDD>=  C220 D106
      ANDD<=  C220 D108
      AND     M222
      OUT     Y040
      MRD
      ANDD>=  C220 D90
      SET     M17
      MRD
      LD      M17
      LDI     M17
      AND     X001
      ANDD>=  C220 K630
      ORB
      ANB
      LD      M222
      LDI     M222
      AND     X005
      ORB
      ANB
      OUT     T14 K10
      MRD
      AND     T14
      AND     M222
      SET     S6
      MRD
      LDD<    C220 D90
      LDI     M14
      ANI     X006
      ORB
      ANB
      ANI     X001
      LD      X023
      ORI     M551
      ANB
      OUT     Y030
      MPP
      AND     Y000
      LD      M222
      LDI     M222
      ANI     M17
      ORB
      ANB
      OUT     M8
8865  LD      M552
      AND     M551
      AND     M528
      LDD>    C220 D36
      LDD>    C220 K300
      AND     X003
      ORB
      ANB
      ANI     M222
      ANI     M223
      ANI     M224
      ANI     M225
      ANI     M226
      ANI     M227
      AND     M228
      SET     M186
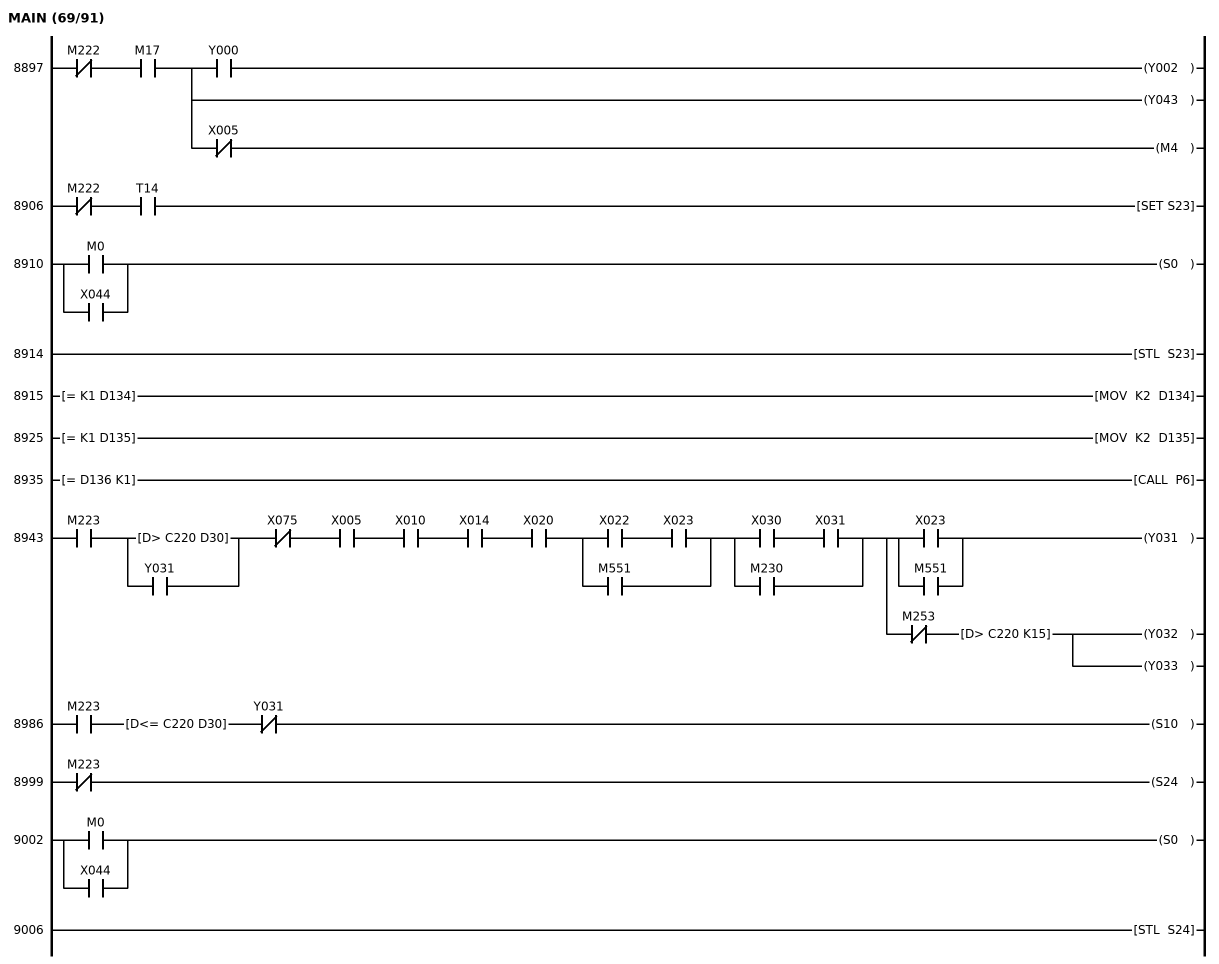
8897  LDI     M222
      AND     M17
      MPS
      AND     Y000
      OUT     Y002
      MPP
      OUT     Y043
      ANI     X005
      OUT     M4
8906  LDI     M222
      AND     T14
      SET     S23
8910  LD      M0
      OR      X044
      OUT     S0
8914  STL     S23
8915  LD=     K1 D134
      MOV     K2 D134
8925  LD=     K1 D135
      MOV     K2 D135
8935  LD=     D136 K1
      CALL    P6
8943  LD      M223
      LDD>    C220 D30
      OR      Y031
      ANB
      ANI     X075
      AND     X005
      AND     X010
      AND     X014
      AND     X020
      LD      X022
      AND     X023
      OR      M551
      ANB
      LD      X030
      AND     X031
      OR      M230
      ANB
      MPS
      LD      X023
      OR      M551
      ANB
      OUT     Y031
      MPP
      ANI     M253
      ANDD>   C220 K15
      OUT     Y032
      OUT     Y033
8986  LD      M223
      ANDD<=  C220 D30
      ANI     Y031
      OUT     S10
8999  LDI     M223
      OUT     S24
9002  LD      M0
      OR      X044
      OUT     S0
9006  STL     S24
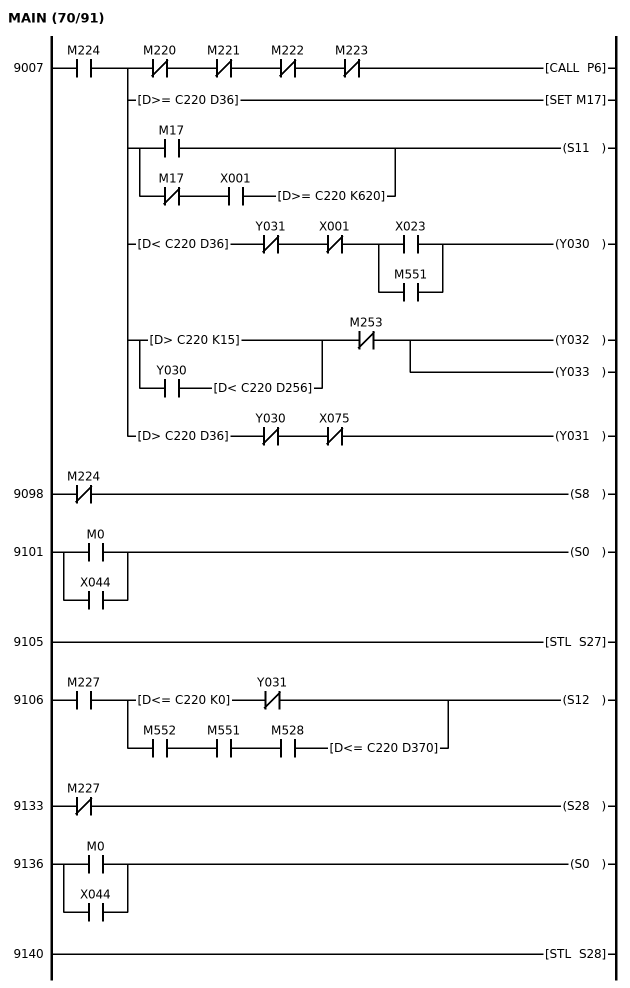
9007  LD      M224
      MPS
      ANI     M220
      ANI     M221
      ANI     M222
      ANI     M223
      CALL    P6
      MRD
      ANDD>=  C220 D36
      SET     M17
      MRD
      LD      M17
      LDI     M17
      AND     X001
      ANDD>=  C220 K620
      ORB
      ANB
      OUT     S11
      MRD
      ANDD<   C220 D36
      ANI     Y031
      ANI     X001
      LD      X023
      OR      M551
      ANB
      OUT     Y030
      MRD
      LDD>    C220 K15
      LD      Y030
      ANDD<   C220 D256
      ORB
      ANB
      ANI     M253
      OUT     Y032
      OUT     Y033
      MPP
      ANDD>   C220 D36
      ANI     Y030
      ANI     X075
      OUT     Y031
9098  LDI     M224
      OUT     S8
9101  LD      M0
      OR      X044
      OUT     S0
9105  STL     S27
9106  LD      M227
      LDD<=   C220 K0
      ANI     Y031
      LD      M552
      AND     M551
      AND     M528
      ANDD<=  C220 D370
      ORB
      ANB
      OUT     S12
9133  LDI     M227
      OUT     S28
9136  LD      M0
      OR      X044
      OUT     S0
9140  STL     S28
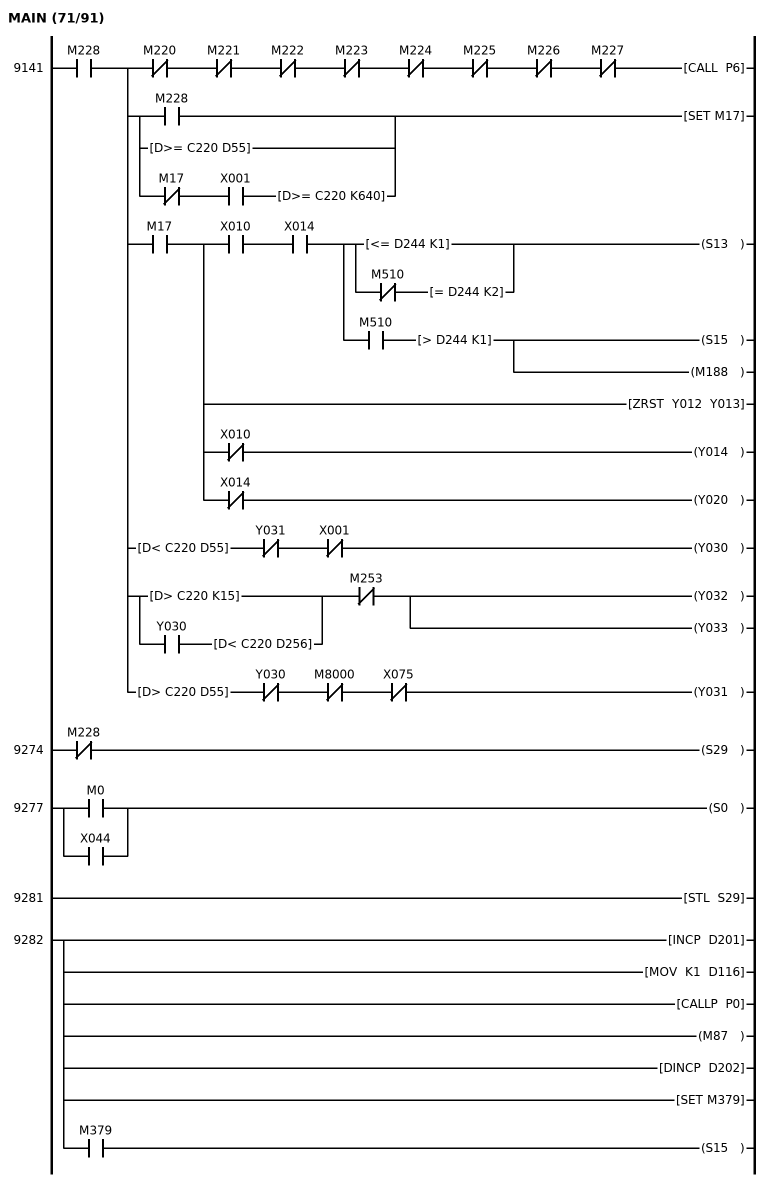
9141  LD      M228
      MPS
      ANI     M220
      ANI     M221
      ANI     M222
      ANI     M223
      ANI     M224
      ANI     M225
      ANI     M226
      ANI     M227
      CALL    P6
      MRD
      LD      M228
      ORD>=   C220 D55
      LDI     M17
      AND     X001
      ANDD>=  C220 K640
      ORB
      ANB
      SET     M17
      MRD
      AND     M17
      MPS
      AND     X010
      AND     X014
      MPS
      LD<=    D244 K1
      LDI     M510
      AND=    D244 K2
      ORB
      ANB
      OUT     S13
      MPP
      AND     M510
      AND>    D244 K1
      OUT     S15
      OUT     M188
      MPP
      ZRST    Y012 Y013
      MPS
      ANI     X010
      OUT     Y014
      MPP
      ANI     X014
      OUT     Y020
      MRD
      ANDD<   C220 D55
      ANI     Y031
      ANI     X001
      OUT     Y030
      MRD
      LDD>    C220 K15
      LD      Y030
      ANDD<   C220 D256
      ORB
      ANB
      ANI     M253
      OUT     Y032
      OUT     Y033
      MPP
      ANDD>   C220 D55
      ANI     Y030
      ANI     M8000
      ANI     X075
      OUT     Y031
9274  LDI     M228
      OUT     S29
9277  LD      M0
      OR      X044
      OUT     S0
9281  STL     S29
9282  INCP    D201
      MOV     K1 D116
      CALLP   P0
      OUT     M87
      DINCP   D202
      SET     M379
      AND     M379
      OUT     S15
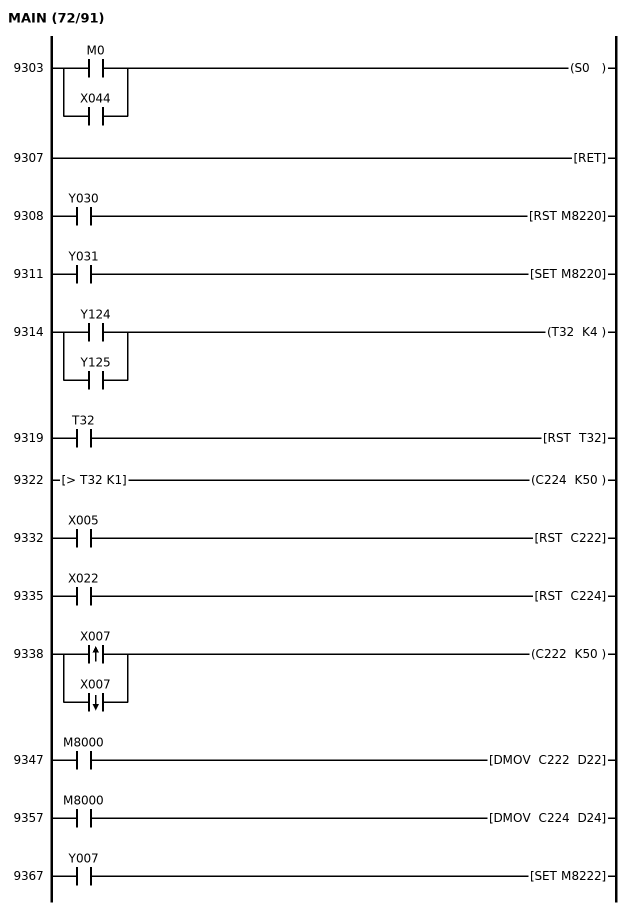
9303  LD      M0
      OR      X044
      OUT     S0
9307  RET
9308  LD      Y030
      RST     M8220
9311  LD      Y031
      SET     M8220
9314  LD      Y124
      OR      Y125
      OUT     T32 K4
9319  LD      T32
      RST     T32
9322  LD>     T32 K1
      OUT     C224 K50
9332  LD      X005
      RST     C222
9335  LD      X022
      RST     C224
9338  LDP     X007
      ORF     X007
      OUT     C222 K50
9347  LD      M8000
      DMOV    C222 D22
9357  LD      M8000
      DMOV    C224 D24
9367  LD      Y007
      SET     M8222
